Staubli VAL3: start.pgx

program start()
begin
  taskCreate "appMain",100,Main()
end
